Fanuc KAREL source: kb00034.KL

-- PROVISIONAL review KL for V1013-1; original PC SHA256 443c43b821ea59e249e2f61ea2c22a01ce6c31957a88cec51e33763ed29b6dff
-- Incomplete behavior may be omitted. Consult companion uncertainty JSON. Do not deploy.
PROGRAM KB00034
%NOLOCKGROUP
BEGIN
  -- UNRESOLVED_PC offsets 5-14; opcodes 3F,75
  -- UNRESOLVED_PC offsets 19-37; opcodes 27,22,22,2A,31
  -- UNRESOLVED_PC offsets 42-46; opcodes 7F
END KB00034
